    rq_activate_all_grippers(True)
    # end: URCap Program Node
  end
  $ 64 "zero_ftsensor()"
  zero_ftsensor()
  $ 65 "EXTT"
  $ 66 "Set GRP_3F_Enable=Off"
  set_standard_digital_out(4, False)
  $ 67 "Set BarcodeTrigger=Off"
  set_standard_digital_out(6, False)
  $ 68 "Set GRP_3F_Decap=Off"
  set_standard_digital_out(3, False)
  $ 69 "Set GRP_3F_Cap=Off"
  set_standard_digital_out(2, False)
  $ 70 "Set GRP_3F_Open=Off"
  set_standard_digital_out(5, False)
  $ 71 "PSE_T≔get_tool_free_pose(dir=[0,0,0.150], move_in_base_frame=True)"
  global PSE_T=get_tool_free_pose(dir=[0,0,0.150], move_in_base_frame=True)
  $ 72 "If is_reachable(Base_const, [PSE_T])"
  if (is_reachable(p[0.0,0.0,0.0,0.0,0.0,0.0], [PSE_T])):
    $ 73 "MoveL"
    $ 74 "PSE_T" "breakAfter"
    movel(PSE_T, a=1.2, v=0.15)
  end
  $ 76 "powder dispensing variable init"
  $ 77 "Start_thread≔ False "
  global Start_thread=  False
  $ 78 "vib_thread≔ False "
  global vib_thread=  False
  $ 79 "QR assignment init"
  $ 80 "d_cc≔0.06"
  global d_cc=0.06
  $ 81 "W_EMPTY≔50.131"
  global W_EMPTY=50.131
  $ 82 "kp≔0.0015"
  global kp=0.0015
  $ 83 "ki≔0.0001"
  global ki=0.0001
  $ 84 "kd≔0.01"
  global kd=0.01
  $ 85 "dt≔0.03"
  global dt=0.03
  $ 86 "Integral_error≔0"
  global Integral_error=0
  $ 87 "current_error≔0"
  global current_error=0
  $ 88 "previous_error≔0"
  global previous_error=0
  $ 89 "tilt_increment≔0"
  global tilt_increment=0
  $ 90 "tilt_angle≔0"
  global tilt_angle=0
  $ 91 "diff≔0"
  global diff=0
  $ 92 "current_pose≔get_actual_tcp_pose()"
  global current_pose= get_actual_tcp_pose ()
  $ 93 "Relative_trans≔p[0, 0, -0.035, 0, 0, 0]"
  global Relative_trans=p[0, 0, -0.035, 0, 0, 0]
  $ 97 "tilt_init_reference()"
  tilt_init_reference()
  $ 98 "switch_spat_M≔ True "
  global switch_spat_M=  True
  $ 99 "switch_spat_S≔ True "
  global switch_spat_S=  True
  $ 100 "switch_spat_F_M≔ True "
  global switch_spat_F_M=  True
  $ 101 "switch_spat_F_S≔ True "
  global switch_spat_F_S=  True
  $ 102 "last_scale≔0"
  global last_scale=0
  $ 775 "Thread_1"
  thread Thread_1():
    while (True):
      $ 776 "If Start_thread≟ True "
      if (Start_thread ==   True  ):
        $ 777 "weight_value≔get_weight()"
        global weight_value=get_weight()
        $ 778 "Wait: 0.1"
        sleep(0.1)
        $ 779 "sync()"
        sync()
      end
      $ 780 "sync()"
      sync()
    end
  end
  threadId_Thread_1 = run Thread_1()
  $ 781 "Thread_2"
  thread Thread_2():
    while (True):
      $ 782 "Loop vib_thread≟ True "
      thread Thread_while_782():
        while (True):
          $ 783 "diff≔target_weight-weight_value"
          global diff=target_weight-weight_value
          $ 784 "If diff>0.02 and spatula≠'spatula_flat_S'"
          global thread_flag_784=0
          thread Thread_if_784():
            $ 786 "Set AO[0]=4.0"
            set_standard_analog_out(0, 0.4)
            thread_flag_784 = 1
          end
          if (diff>0.02  and  spatula != "spatula_flat_S"):
            global thread_handler_784=run Thread_if_784()
            while (thread_flag_784 == 0):
              if not(diff>0.02  and  spatula != "spatula_flat_S"):
                kill thread_handler_784
                thread_flag_784 = 2
              else:
                sync()
              end
            end
          else:
            thread_flag_784 = 2
          end
          if (thread_flag_784 == 2):
            $ 787 "ElseIf diff>0.02 and spatula≟'spatula_flat_S'"
            if (diff>0.02 and spatula == "spatula_flat_S"):
              $ 788 "vibration_3()"
              vibration_3()
            else:
              $ 789 "ElseIf diff≤0.03"
              global thread_flag_789=0
              thread Thread_if_789():
                $ 790 "vibration_2()"
                vibration_2()
                thread_flag_789 = 1
              end
              if (diff <= 0.03):
                global thread_handler_789=run Thread_if_789()
                while (thread_flag_789 == 0):
                  if not(diff <= 0.03):
                    kill thread_handler_789
                    thread_flag_789 = 2
                  else:
                    sync()
                  end
                end
              else:
                thread_flag_789 = 2
              end
              if (thread_flag_789 == 2):
                $ 795 "Else" "noBreak"
                $ 796 "Set AO[0]=0.0"
                set_standard_analog_out(0, 0.0)
              end
            end
          end
        end
      end
      if (vib_thread ==   True  ):
        global thread_handler_782=run Thread_while_782()
        while (vib_thread ==   True  ):
          sync()
        end
        kill thread_handler_782
      end
      $ 797 "sync()"
      sync()
    end
  end
  threadId_Thread_2 = run Thread_2()
  while (True):
    $ 103 "Robot Program"
    $ 104 "MAIN"
    $ 105 "command_manager(external_control='uGO', cond_suspend=(ITM_Manipulated and AMR_AtTarget and AMR_Charging and AMR_Battery<40), cond_unsuspend=(AMR_Battery≟60))"
    command_manager(external_control="uGO", cond_suspend=(ITM_Manipulated  and  AMR_AtTarget  and  AMR_Charging  and  AMR_Battery<40), cond_unsuspend=(AMR_Battery == 60))
    $ 106 "log_state(STATE_Info)"
    log_state(STATE_Info)
    $ 107 "Switch STATE"
    switch_1 = STATE
    $ 108 "Case 1"
    if (1 == switch_1):
      $ 109 "Stopping"
      $ 110 "STATE_Info≔'Stopping'"
      global STATE_Info="Stopping"
      $ 111 "end_freedrive_mode()"
      end_freedrive_mode()
      $ 112 "Set"
      set_tcp(p[0.0,0.0,0.161,3.1415,0.0,0.0])
      $ 113 "PSE_T≔get_tool_free_pose(dir=[0,0,0.150], move_in_base_frame=True)"
      global PSE_T=get_tool_free_pose(dir=[0,0,0.150], move_in_base_frame=True)
      $ 114 "If is_reachable(Base_const, [PSE_T])"
      if (is_reachable(p[0.0,0.0,0.0,0.0,0.0,0.0], [PSE_T])):
        $ 115 "MoveL"
        $ 116 "PSE_T" "breakAfter"
        movel(PSE_T, a=1.2, v=0.15)
      end
      $ 117 "do_transition(keep_rxry=OBJ_Picked, r=0)"
      do_transition(keep_rxry=OBJ_Picked, r=0)
      $ 126 "Call Sub_AMR_MiR_V3"
      Sub_AMR_MiR_V3()
      $ 127 "If stopping() and AMR_Done"
      if (stopping()  and  AMR_Done):
        $ 128 "STATE≔2"
        global STATE=2
        $ 129 "ugo_update_outputs()"
        ugo_update_outputs()
      end
    elif (2 == switch_1):
      $ 130 "Case 2"
      $ 131 "Stopped"
      $ 132 "STATE_Info≔'Stopped'"
      global STATE_Info="Stopped"
      $ 133 "Call Sub_AMR_MiR_V3"
      Sub_AMR_MiR_V3()
      $ 134 "If CMD_Reset  or PB_Start"
      if (CMD_Reset   or  get_standard_digital_in(0)):
        $ 135 "STATE≔3"
        global STATE=3
        $ 136 "ugo_update_outputs()"
        ugo_update_outputs()
      end
    elif (3 == switch_1):
      $ 137 "Case 3"
      $ 138 " Resetting"
      $ 139 "STATE_Info≔'Resetting'"
      global STATE_Info="Resetting"
      $ 140 "uML"
      $ 141 "reset_error()"
      reset_error()
      $ 142 "reset_warning()"
      reset_warning()
      $ 143 "PROCESS_Step≔0"
      global PROCESS_Step=0
      $ 144 "PROCESS_Info≔''"
      global PROCESS_Info=""
      $ 145 "ARM_Referenced≔ False "
      global ARM_Referenced=  False
      $ 146 "WRK_Done≔ False "
      global WRK_Done=  False
      $ 147 "ITM_Prepared≔ False "
      global ITM_Prepared=  False
      $ 148 "ITM_Manipulated≔ False "
      global ITM_Manipulated=  False
      $ 149 "STP≔0"
      global STP=0
      $ 150 "Action≔0"
      global Action=0
      $ 151 "Action_Info≔''"
      global Action_Info=""
      $ 152 "ITM_ID≔0"
      global ITM_ID=0
      $ 153 "JIG≔0"
      global JIG=0
      $ 154 "JIG_Slot≔0"
      global JIG_Slot=0
      $ 155 "Task_info≔''"
      global Task_info=""
      $ 156 "Set"
      set_tcp(p[0.0,0.0,0.161,3.1415,0.0,0.0])
      $ 157 "App"
      $ 158 "'ADD APPLICATION SPECIFIC COMMANDS'"
      # 'ADD APPLICATION SPECIFIC COMMANDS'
      $ 159 "OBJ_Type≔0"
      global OBJ_Type=0
      $ 160 "OBJ_Nbr≔0"
      global OBJ_Nbr=0
      $ 161 "If CNT_Rack_Output≥50"
      if (CNT_Rack_Output >= 50):
        $ 162 "CNT_Rack_Output≔0"
        global CNT_Rack_Output=0
      end
      $ 163 "TASK≔struct(ID=0, NAVI=struct(target=0, footprint=0, protectiveOff=0, dock=0), WORK=struct(ITM_ID_Src=0, JIG_ID_Src=0, OBJ_Nbr_Src=0, ACT_Src=0, ITM_ID_Tgt=0, JIG_ID_Tgt=0, OBJ_Nbr_Tgt=0, ACT_Tgt=0, OBJ_Type=0))"
      global TASK=struct(ID=0, NAVI=struct(target=0, footprint=0, protectiveOff=0, dock=0), WORK=struct(ITM_ID_Src=0, JIG_ID_Src=0, OBJ_Nbr_Src=0, ACT_Src=0, ITM_ID_Tgt=0, JIG_ID_Tgt=0, OBJ_Nbr_Tgt=0, ACT_Tgt=0, OBJ_Type=0))
      $ 164 "Call Sub_AMR_MiR_V3"
      Sub_AMR_MiR_V3()
      $ 165 "If resetting() and AMR_Done"
      if (resetting()  and  AMR_Done):
        $ 166 "STATE≔4"
        global STATE=4
        $ 167 "ugo_update_outputs()"
        ugo_update_outputs()
      end
    elif (4 == switch_1):
      $ 168 "Case 4"
      $ 169 "Idle"
      $ 170 "STATE_Info≔'Idle'"
      global STATE_Info="Idle"
      $ 171 "If CMD_Start"
      if (CMD_Start):
        $ 172 "STATE≔5"
        global STATE=5
        $ 173 "ugo_update_outputs()"
        ugo_update_outputs()
      end
    elif (5 == switch_1):
      $ 174 "Case 5"
      $ 175 "Starting"
      $ 176 "STATE_Info≔'Starting'"
      global STATE_Info="Starting"
      $ 177 "'ADD COMMANDS WHAT TO START WITH'"
      # 'ADD COMMANDS WHAT TO START WITH'
      $ 178 "Call Sub_AMR_MiR_V3"
      Sub_AMR_MiR_V3()
      $ 179 "get ugo data"
      $ 180 "Assign Tasks"
      $ 181 "TASK.ID = ugo_get_task()"
      TASK.ID = ugo_get_task()
      $ 182 "If TASK.ID≟1"
      if (TASK.ID == 1):
        $ 183 "Task_info≔'Charge'"
        global Task_info="Charge"
        $ 184 "Parameters"
        $ 185 "AMR_PosTarget≔1"
        global AMR_PosTarget=1
      else:
        $ 186 "ElseIf TASK.ID≟9"
        if (TASK.ID == 9):
          $ 187 "'Pick Sarstedt Rack from Variable source'"
          # 'Pick Sarstedt Rack from Variable source'
          $ 188 "Task_info≔'Navigate to Target'"
          global Task_info="Navigate to Target"
          $ 189 "Parameters"
          $ 190 "AMR_PosTarget≔UGO.read_input('00','ITM_ID')"
          global AMR_PosTarget=UGO.read_input("00","ITM_ID")
        else:
          $ 191 "ElseIf TASK.ID≟49"
          if (TASK.ID == 49):
            $ 192 "Task_info≔'Pick Containers'"
            global Task_info="Pick Containers"
            $ 193 "Parameters"
            $ 194 "ITM_ID≔1"
            global ITM_ID=1
            $ 195 "OBJ_Type≔6"
            global OBJ_Type=6
            $ 196 "JIG≔15"
            global JIG=15
            $ 197 "AMR_PosTarget≔3"
            global AMR_PosTarget=3
          else:
            $ 198 "ElseIf TASK.ID≟50"
            if (TASK.ID == 50):
              $ 199 "Task_info≔'Decap Containers'"
              global Task_info="Decap Containers"
              $ 200 "Parameters"
              $ 201 "ITM_ID≔1"
              global ITM_ID=1
              $ 202 "OBJ_Type≔6"
              global OBJ_Type=6
              $ 203 "JIG≔16"
              global JIG=16
              $ 204 "AMR_PosTarget≔5"
              global AMR_PosTarget=5
            else:
              $ 205 "ElseIf TASK.ID≟51"
              if (TASK.ID == 51):
                $ 206 "Task_info≔'Detect Spatula and transfer powder'"
                global Task_info="Detect Spatula and transfer powder"
                $ 207 "Parameters"
                $ 208 "ITM_ID≔1"
                global ITM_ID=1
                $ 209 "target_weight≔(UGO.read_input('00','Target_weight'))/1000"
                global target_weight=(UGO.read_input("00","Target_weight"))/1000
                $ 210 "OBJ_Type≔8"
                global OBJ_Type=8
                $ 211 "JIG≔16"
                global JIG=16
                $ 212 "AMR_PosTarget≔5"
                global AMR_PosTarget=5
              else:
                $ 213 "ElseIf TASK.ID≟52"
                if (TASK.ID == 52):
                  $ 214 "Task_info≔'Pick Powder'"
                  global Task_info="Pick Powder"
                  $ 215 "Parameters"
                  $ 216 "ITM_ID≔1"
                  global ITM_ID=1
                  $ 217 "OBJ_Type≔6"
                  global OBJ_Type=6
                  $ 218 "JIG≔15"
                  global JIG=15
                  $ 219 "AMR_PosTarget≔3"
                  global AMR_PosTarget=3
                else:
                  $ 220 "ElseIf TASK.ID≟53"
                  if (TASK.ID == 53):
                    $ 221 "Task_info≔'Decap Powder'"
                    global Task_info="Decap Powder"
                    $ 222 "Parameters"
                    $ 223 "ITM_ID≔1"
                    global ITM_ID=1
                    $ 224 "OBJ_Type≔6"
                    global OBJ_Type=6
                    $ 225 "JIG≔1"
                    global JIG=1
                    $ 226 "AMR_PosTarget≔5"
                    global AMR_PosTarget=5
                  else:
                    $ 227 "ElseIf TASK.ID≟54"
                    if (TASK.ID == 54):
                      $ 228 "Task_info≔'Empty and swap Powder container'"
                      global Task_info="Empty and swap Powder container"
                      $ 237 "Parameters"
                      $ 238 "ITM_ID≔1"
                      global ITM_ID=1
                      $ 240 "W_now≔(UGO.read_input('00','Container_weight'))/1000"
                      global W_now=(UGO.read_input("00","Container_weight"))/1000
                      $ 241 "Pow_name≔(UGO.read_input('00','Powder_name'))"
                      global Pow_name=(UGO.read_input("00","Powder_name"))
                      $ 242 "scooping_init()"
                      scooping_init()
                      $ 243 "target_weight≔W_now-W_EMPTY-(0.002*W_FULL)"
                      global target_weight=W_now-W_EMPTY-(0.002*W_FULL)
                      $ 244 "OBJ_Type≔6"
                      global OBJ_Type=6
                      $ 245 "JIG≔17"
                      global JIG=17
                      $ 246 "AMR_PosTarget≔5"
                      global AMR_PosTarget=5
                    else:
                      $ 247 "ElseIf TASK.ID≟55"
                      if (TASK.ID == 55):
                        $ 248 "Task_info≔'Place Powder'"
                        global Task_info="Place Powder"
                        $ 249 "Parameters"
                        $ 250 "ITM_ID≔1"
                        global ITM_ID=1
                        $ 251 "OBJ_Type≔6"
                        global OBJ_Type=6
                        $ 252 "JIG≔21"
                        global JIG=21
                        $ 253 "AMR_PosTarget≔5"
                        global AMR_PosTarget=5
                      else:
                        $ 254 "ElseIf TASK.ID≟56"
                        if (TASK.ID == 56):
                          $ 255 "Task_info≔'Dose Powder'"
                          global Task_info="Dose Powder"
                          $ 256 "Parameters"
                          $ 257 "ITM_ID≔1"
                          global ITM_ID=1
                          $ 258 "target_weight≔(UGO.read_input('00','Target_weight'))/1000"
                          global target_weight=(UGO.read_input("00","Target_weight"))/1000
                          $ 259 "W_now≔(UGO.read_input('00','Container_weight'))/1000"
                          global W_now=(UGO.read_input("00","Container_weight"))/1000
                          $ 261 "Pow_name≔(UGO.read_input('00','Powder_name'))"
                          global Pow_name=(UGO.read_input("00","Powder_name"))
                          $ 262 "OBJ_Type≔6"
                          global OBJ_Type=6
                          $ 263 "JIG≔17"
                          global JIG=17
                          $ 264 "AMR_PosTarget≔5"
                          global AMR_PosTarget=5
                        else:
                          $ 265 "ElseIf TASK.ID≟57"
                          if (TASK.ID == 57):
                            $ 266 "Task_info≔'Recipe Powder dosing'"
                            global Task_info="Recipe Powder dosing"
                            $ 267 "Parameters"
                            $ 268 "ITM_ID≔1"
                            global ITM_ID=1
                            $ 269 "Pow_A≔(UGO.read_input('00','PowderA'))"
                            global Pow_A=(UGO.read_input("00","PowderA"))
                            $ 270 "Pow_B≔(UGO.read_input('00','PowderB'))"
                            global Pow_B=(UGO.read_input("00","PowderB"))
                            $ 271 "Pow_C≔(UGO.read_input('00','PowderC'))"
                            global Pow_C=(UGO.read_input("00","PowderC"))
                            $ 272 "Total_weight≔(UGO.read_input('00','Total_weight'))/1000"
                            global Total_weight=(UGO.read_input("00","Total_weight"))/1000
                            $ 273 "Pow_A_percent≔(UGO.read_input('00','PowderA_percentage'))/100"
                            global Pow_A_percent=(UGO.read_input("00","PowderA_percentage"))/100
                            $ 274 "Pow_B_percent≔(UGO.read_input('00','PowderB_percentage'))/100"
                            global Pow_B_percent=(UGO.read_input("00","PowderB_percentage"))/100
                            $ 275 "Pow_C_percent≔(UGO.read_input('00','PowderC_percentage'))/100"
                            global Pow_C_percent=(UGO.read_input("00","PowderC_percentage"))/100
                            $ 276 "OBJ_Type≔6"
                            global OBJ_Type=6
                            $ 277 "JIG≔17"
                            global JIG=17
                            $ 278 "AMR_PosTarget≔5"
                            global AMR_PosTarget=5
                          else:
                            $ 279 "ElseIf TASK.ID≟58"
                            if (TASK.ID == 58):
                              $ 280 "Task_info≔'Pick Powder containers'"
                              global Task_info="Pick Powder containers"
                              $ 281 "Parameters"
                              $ 282 "ITM_ID≔1"
                              global ITM_ID=1
                              $ 283 "OBJ_Type≔6"
                              global OBJ_Type=6
                              $ 284 "JIG≔15"
                              global JIG=15
                              $ 285 "AMR_PosTarget≔3"
                              global AMR_PosTarget=3
                            else:
                              $ 286 "Else" "noBreak"
                              $ 287 "set_error(ERROR_WRONG_ORDER)"
                              set_error(ERROR_WRONG_ORDER)
                            end
                          end
                        end
                      end
                    end
                  end
                end
              end
            end
          end
        end
      end
      $ 288 "test ugo"
      $ 289 "Wait: 0.2"
      sleep(0.2)
      $ 290 "ugo_update_outputs()"
      ugo_update_outputs()
      $ 291 "If starting() and AMR_Done"
      if (starting()  and  AMR_Done):
        $ 292 "log_message(Task_info, 'New Task: ')"
        log_message(Task_info, "New Task: ")
        $ 293 "log_message(to_str(TASK.ID), 'Task_ID: ')"
        log_message(to_str(TASK.ID), "Task_ID: ")
        $ 294 "do_transition(keep_rxry=OBJ_Picked)"
        do_transition(keep_rxry=OBJ_Picked)
        $ 295 "STATE≔6"
        global STATE=6
        $ 296 "ugo_update_outputs()"
        ugo_update_outputs()
      end
    elif (6 == switch_1):
      $ 297 "Case 6"
      $ 298 "Execute"
      $ 299 "STATE_Info≔'Execute'"
      global STATE_Info="Execute"
      $ 300 "If  not CMD_Hold and not CMD_Suspend"
      global thread_flag_300=0
      thread Thread_if_300():
        $ 301 "Switch PROCESS_Step"
        switch_2 = PROCESS_Step
        $ 302 "Case 0"
        if (0 == switch_2):
          $ 303 "PROCESS_Info≔'process control'"
          global PROCESS_Info="process control"
          $ 304 "log_process(PROCESS_Info)"
          log_process(PROCESS_Info)
          $ 305 "process control"
          $ 306 "If  not AMR_AtTarget"
          if (  not  AMR_AtTarget):
            $ 307 "PROCESS_Step≔1"
            global PROCESS_Step=1
          else:
            $ 308 "ElseIf (( not ITM_Prepared and  not WRK_Done) or (ITM_Prepared and WRK_Done))"
            if (((  not  ITM_Prepared  and    not  WRK_Done)  or  (ITM_Prepared  and  WRK_Done))):
              $ 309 "PROCESS_Step≔2"
              global PROCESS_Step=2
            else:
              $ 310 "ElseIf  not WRK_Done"
              if (  not  WRK_Done):
                $ 311 "PROCESS_Step≔3"
                global PROCESS_Step=3
              else:
                $ 312 "Else" "noBreak"
                $ 313 "task finished"
                $ 314 "PROCESS_Info≔''"
                global PROCESS_Info=""
                $ 315 "STATE≔7"
                global STATE=7
                $ 316 "ugo_update_outputs()"
                ugo_update_outputs()
              end
            end
          end
        elif (1 == switch_2):
          $ 317 "Case 1"
          $ 318 "navigate"
          $ 319 "'MOVING THE uML'"
          # 'MOVING THE uML'
          $ 320 "PROCESS_Info≔'move to target'"
          global PROCESS_Info="move to target"
          $ 321 "log_process(PROCESS_Info)"
          log_process(PROCESS_Info)
          $ 322 "If TASK.ID≟1"
          if (TASK.ID == 1):
            $ 323 "Action≔51"
            global Action=51
          else:
            $ 324 "Else" "noBreak"
            $ 325 "Action≔52"
            global Action=52
          end
          $ 326 "Call Sub_AMR_MiR_V3"
          Sub_AMR_MiR_V3()
          $ 327 "If AMR_Done"
          if (AMR_Done):
            $ 328 "PROCESS_Step≔0"
            global PROCESS_Step=0
          end
        elif (2 == switch_2):
          $ 329 "Case 2"
          $ 330 "prepare"
          $ 331 "'THINGS THAT HAVE TO BE DONE ONCE IN A SEQUENCE,WORKFLOW'"
          # 'THINGS THAT HAVE TO BE DONE ONCE IN A SEQUENCE,WORKFLOW'
          $ 332 "PROCESS_Info≔'prepare for work'"
          global PROCESS_Info="prepare for work"
          $ 333 "log_process(PROCESS_Info)"
          log_process(PROCESS_Info)
          $ 334 "If TASK.WORK.ITM_ID_Src>1"
          if (TASK.WORK.ITM_ID_Src>1):
            $ 335 "ITM_ID≔TASK.WORK.ITM_ID_Src"
            global ITM_ID=TASK.WORK.ITM_ID_Src
          else:
            $ 336 "ElseIf TASK.WORK.ITM_ID_Tgt>1"
            if (TASK.WORK.ITM_ID_Tgt>1):
              $ 337 "ITM_ID≔TASK.WORK.ITM_ID_Tgt"
              global ITM_ID=TASK.WORK.ITM_ID_Tgt
            end
          end
          $ 338 "If  not ARM_Referenced and (ITM_ID≠0)"
          if (  not  ARM_Referenced  and  (ITM_ID != 0)):
            $ 339 "STP≔1"
            global STP=1
          else:
            $ 340 "ElseIf ARM_Referenced or (ITM_ID≟0)"
            if (ARM_Referenced  or  (ITM_ID == 0)):
              $ 341 "STP≔2"
              global STP=2
            end
          end
          $ 342 "Switch STP"
          switch_3 = STP
          $ 343 "Case 1"
          if (1 == switch_3):
            $ 344 "reference"
            $ 345 "STP_Info≔'reference at target position'"
            global STP_Info="reference at target position"
            $ 346 "log_step(STP_Info)"
            log_step(STP_Info)
            $ 347 "If ITM_ID≟1"
            if (ITM_ID == 1):
              $ 348 "CAM_Done≔ True "
              global CAM_Done=  True
            else:
              $ 349 "Else" "noBreak"
              $ 350 "Action≔131"
              global Action=131
              $ 351 "Call Sub_Vision_V18"
              Sub_Vision_V18()
            end
            $ 353 "If CAM_Done and  not ERROR.FLAG"
            if (CAM_Done  and    not  ERROR.FLAG):
              $ 354 "log_step('ARM referenced')"
              log_step("ARM referenced")
              $ 355 "ARM_Referenced≔ True "
              global ARM_Referenced=  True
            end
          elif (2 == switch_3):
            $ 356 "Case 2"
            $ 357 "manipulate"
            $ 358 "STP_Info≔'manipulate item'"
            global STP_Info="manipulate item"
            $ 359 "log_step(STP_Info)"
            log_step(STP_Info)
            $ 360 "'In case pressing button is needed'"
            # 'In case pressing button is needed'
            $ 361 "If found_in_list(ITM_ID, ITM_ID_List)"
            if (found_in_list(ITM_ID, ITM_ID_List)):
              $ 362 "Switch ITM_ID"
              switch_4 = ITM_ID
              $ 363 "Case 0"
              if (0 == switch_4):
                $ 364 "ITM_Manipulated≔ not ITM_Manipulated"
                global ITM_Manipulated=  not  ITM_Manipulated
              elif (1 == switch_4):
                $ 365 "Case 1"
                $ 366 "ITM_Manipulated≔ not ITM_Manipulated"
                global ITM_Manipulated=  not  ITM_Manipulated
              elif (2 == switch_4):
                $ 367 "Case 2"
              else:
                $ 377 "Default Case"
                $ 378 "ITM_Manipulated≔ not ITM_Manipulated"
                global ITM_Manipulated=  not  ITM_Manipulated
              end
            end
          end
          $ 379 "ITM_Prepared≔(ITM_Manipulated or  not found_in_list(ITM_ID, ITM_ID_List)) and (ARM_Referenced or ITM_ID≟0) and  not WRK_Done"
          global ITM_Prepared=(ITM_Manipulated  or    not  found_in_list(ITM_ID, ITM_ID_List))  and  (ARM_Referenced  or  ITM_ID == 0)  and    not  WRK_Done
          $ 380 "STP≔0"
          global STP=0
          $ 381 "STP_Info≔''"
          global STP_Info=""
          $ 382 "PROCESS_Step≔0"
          global PROCESS_Step=0
        elif (3 == switch_2):
          $ 383 "Case 3"
          $ 384 "work"
          $ 385 "'ADD EVERY MACHINE, OBJECT, STATION TO WORK ON'"
          # 'ADD EVERY MACHINE, OBJECT, STATION TO WORK ON'
          $ 386 "Switch ITM_ID"
          switch_3 = ITM_ID
          $ 387 "Case 1"
          if (1 == switch_3):
            $ 388 "uLM"
            $ 389 "If TASK.ID≟12"
            if (TASK.ID == 12):
              $ 390 "fill racks"
              $ 391 "Action≔151"
              global Action=151
              $ 392 "Call Sub_Vision_V18"
              Sub_Vision_V18()
              $ 393 "If  not ERROR.FLAG"
              if (  not  ERROR.FLAG):
                $ 394 "Actions for the task"
                $ 395 "Action≔1"
                global Action=1
                $ 396 "JIG≔2"
                global JIG=2
                $ 397 "JIG_Slot≔CAM_Result[0]"
                global JIG_Slot=CAM_Result[0]
                $ 398 "OBJ_Nbr≔CAM_Result[0]"
                global OBJ_Nbr=CAM_Result[0]
                $ 399 "OBJ_Type≔2"
                global OBJ_Type=2
                $ 400 "Call Sub_Action_V4"
                Sub_Action_V4()
                $ 401 "If OBJ_Picked"
                if (OBJ_Picked):
                  $ 402 "CAM_Result.remove(0)"
                  CAM_Result.remove(0)
                  $ 403 "PRC_TubCounter≔PRC_TubCounter+1"
                  global PRC_TubCounter=PRC_TubCounter+1
                  $ 404 "If PRC_TubCounter%4≟0"
                  if (PRC_TubCounter%4 == 0):
                    $ 405 "JIG_Slot≔4"
                    global JIG_Slot=4
                  else:
                    $ 406 "Else" "noBreak"
                    $ 407 "JIG_Slot≔PRC_TubCounter%4"
                    global JIG_Slot=PRC_TubCounter%4
                  end
                  $ 408 "OBJ_Nbr≔ceil(PRC_TubCounter/4)"
                  global OBJ_Nbr=ceil(PRC_TubCounter/4)
                  $ 409 "Action≔2"
                  global Action=2
                  $ 410 "JIG≔4"
                  global JIG=4
                  $ 411 "Call Sub_Action_V4"
                  Sub_Action_V4()
                  $ 412 "Action≔151"
                  global Action=151
                  $ 413 "Call Sub_Vision_V18"
                  Sub_Vision_V18()
                end
              end
              $ 414 "If (CAM_Captures≥CAM_PRM_Retries) or (PRC_TubCounter≥32)"
              if ((CAM_Captures >= CAM_PRM_Retries)  or  (PRC_TubCounter >= 32)):
                $ 415 "PROCESS_Step≔0"
                global PROCESS_Step=0
                $ 416 "WRK_Done≔ True "
                global WRK_Done=  True
              end
            else:
              $ 417 "ElseIf TASK.ID≟49"
              if (TASK.ID == 49):
                $ 418 "Pick Powder container"
                $ 419 "Action≔131"
                global Action=131
                $ 420 "Call Sub_Vision_V18"
                Sub_Vision_V18()
                $ 421 "Action≔35"
                global Action=35
                $ 422 "Call Sub_Action_V4"
                Sub_Action_V4()
                $ 423 "PROCESS_Step≔0"
                global PROCESS_Step=0
                $ 424 "WRK_Done≔ True "
                global WRK_Done=  True
              else:
                $ 425 "ElseIf TASK.ID≟50"
                if (TASK.ID == 50):
                  $ 426 "Decap containers"
                  $ 427 "Action≔36"
                  global Action=36
                  $ 428 "Call Sub_Action_V4"
                  Sub_Action_V4()
                  $ 429 "PROCESS_Step≔0"
                  global PROCESS_Step=0
                  $ 430 "WRK_Done≔ True "
                  global WRK_Done=  True
                else:
                  $ 431 "ElseIf TASK.ID≟51"
                  if (TASK.ID == 51):
                    $ 432 "Detect Spatula and transfer powder"
                    $ 433 "Action≔131"
                    global Action=131
                    $ 434 "Call Sub_Vision_V18"
                    Sub_Vision_V18()
                    $ 435 "Action≔37"
                    global Action=37
                    $ 436 "Call Sub_Action_V4"
                    Sub_Action_V4()
                    $ 437 "PROCESS_Step≔0"
                    global PROCESS_Step=0
                    $ 438 "WRK_Done≔ True "
                    global WRK_Done=  True
                  else:
                    $ 439 "ElseIf TASK.ID≟52"
                    if (TASK.ID == 52):
                      $ 440 "Pick Powder container"
                      $ 441 "Action≔131"
                      global Action=131
                      $ 442 "Call Sub_Vision_V18"
                      Sub_Vision_V18()
                      $ 443 "Action≔39"
                      global Action=39
                      $ 444 "Call Sub_Action_V4"
                      Sub_Action_V4()
                      $ 445 "PROCESS_Step≔0"
                      global PROCESS_Step=0
                      $ 446 "WRK_Done≔ True "
                      global WRK_Done=  True
                    else:
                      $ 447 "ElseIf TASK.ID≟53"
                      if (TASK.ID == 53):
                        $ 448 "Decap containerA"
                        $ 449 "Action≔40"
                        global Action=40
                        $ 450 "Call Sub_Action_V4"
                        Sub_Action_V4()
                        $ 451 "PROCESS_Step≔0"
                        global PROCESS_Step=0
                        $ 452 "WRK_Done≔ True "
                        global WRK_Done=  True
                      else:
                        $ 453 "ElseIf TASK.ID≟55"
                        if (TASK.ID == 55):
                          $ 454 "Place Powder"
                          $ 455 "Action≔131"
                          global Action=131
                          $ 456 "Call Sub_Vision_V18"
                          Sub_Vision_V18()
                          $ 457 "Action≔41"
                          global Action=41
                          $ 458 "Call Sub_Action_V4"
                          Sub_Action_V4()
                          $ 459 "PROCESS_Step≔0"
                          global PROCESS_Step=0
                          $ 460 "WRK_Done≔ True "
                          global WRK_Done=  True
                        else:
                          $ 461 "ElseIf TASK.ID≟54"
                          if (TASK.ID == 54):
                            $ 462 "Empty and swap container"
                            $ 463 "Action≔131"
                            global Action=131
                            $ 464 "Call Sub_Vision_V18"
                            Sub_Vision_V18()
                            $ 465 "Action≔42"
                            global Action=42
                            $ 466 "Call Sub_Action_V4"
                            Sub_Action_V4()
                            $ 467 "PROCESS_Step≔0"
                            global PROCESS_Step=0
                            $ 468 "WRK_Done≔ True "
                            global WRK_Done=  True
                          else:
                            $ 469 "ElseIf TASK.ID≟56"
                            if (TASK.ID == 56):
                              $ 470 "Dispense Powder"
                              $ 471 "Action≔131"
                              global Action=131
                              $ 472 "Call Sub_Vision_V18"
                              Sub_Vision_V18()
                              $ 473 "Action≔43"
                              global Action=43
                              $ 474 "Call Sub_Action_V4"
                              Sub_Action_V4()
                              $ 475 "PROCESS_Step≔0"
                              global PROCESS_Step=0
                              $ 476 "WRK_Done≔ True "
                              global WRK_Done=  True
                            else:
                              $ 477 "ElseIf TASK.ID≟57"
                              if (TASK.ID == 57):
                                $ 478 "Recipe Dosing"
                                $ 479 "Action≔48"
                                global Action=48
                                $ 480 "Call Sub_Action_V4"
                                Sub_Action_V4()
                                $ 481 "recipe_init(Pow_A, Pow_B, Pow_C, Total_weight, Pow_A_percent, Pow_B_percent, Pow_C_percent)"
                                recipe_init(Pow_A, Pow_B, Pow_C, Total_weight, Pow_A_percent, Pow_B_percent, Pow_C_percent)
                                $ 482 "Loop recipe_next()≟ True "
                                while (recipe_next() ==   True  ):
                                  $ 483 "Action≔44"
                                  global Action=44
                                  $ 484 "Call Sub_Action_V4"
                                  Sub_Action_V4()
                                  $ 485 "JIG≔21"
                                  global JIG=21
                                  $ 486 "Action≔131"
                                  global Action=131
                                  $ 487 "Call Sub_Vision_V18"
                                  Sub_Vision_V18()
                                  $ 488 "Action≔45"
                                  global Action=45
                                  $ 489 "Call Sub_Action_V4"
                                  Sub_Action_V4()
                                  $ 490 "dosing_start()"
                                  dosing_start()
                                  $ 491 "JIG≔17"
                                  global JIG=17
                                  $ 492 "Action≔131"
                                  global Action=131
                                  $ 493 "Call Sub_Vision_V18"
                                  Sub_Vision_V18()
                                  $ 494 "Action≔46"
                                  global Action=46
                                  $ 495 "Call Sub_Action_V4"
                                  Sub_Action_V4()
                                  $ 496 "dosing_end()"
                                  dosing_end()
                                end
                                $ 497 "PROCESS_Step≔0"
                                global PROCESS_Step=0
                                $ 498 "WRK_Done≔ True "
                                global WRK_Done=  True
                              else:
                                $ 499 "ElseIf TASK.ID≟58"
                                if (TASK.ID == 58):
                                  $ 500 "Pick Powder containers"
                                  $ 501 "Num_cont_picked≔0"
                                  global Num_cont_picked=0
                                  $ 502 "powder_position≔'Position1'"
                                  global powder_position="Position1"
                                  $ 503 "Loop Num_cont_picked<3"
                                  while (Num_cont_picked<3):
                                    $ 504 "Action≔131"
                                    global Action=131
                                    $ 505 "Call Sub_Vision_V18"
                                    Sub_Vision_V18()
                                    $ 506 "Action≔47"
                                    global Action=47
                                    $ 507 "Call Sub_Action_V4"
                                    Sub_Action_V4()
                                  end
                                  $ 508 "PROCESS_Step≔0"
                                  global PROCESS_Step=0
                                  $ 509 "WRK_Done≔ True "
                                  global WRK_Done=  True
                                end
                              end
                            end
                          end
                        end
                      end
                    end
                  end
                end
              end
            end
          elif (2 == switch_3):
            $ 510 "Case 2"
          elif (5 == switch_3):
            $ 552 "Case 5"
          elif (20 == switch_3):
            $ 560 "Case 20"
          elif (43 == switch_3):
            $ 622 "Case 43"
          else:
            $ 630 "Default Case"
            $ 631 "WRK_Done≔ True "
            global WRK_Done=  True
            $ 632 "PROCESS_Step≔0"
            global PROCESS_Step=0
          end
        end
        thread_flag_300 = 1
      end
      if (  not  CMD_Hold and not CMD_Suspend):
        global thread_handler_300=run Thread_if_300()
        while (thread_flag_300 == 0):
          if not(  not  CMD_Hold and not CMD_Suspend):
            kill thread_handler_300
            thread_flag_300 = 2
          else:
            sync()
          end
        end
      else:
        thread_flag_300 = 2
      end
      $ 633 "If CMD_Hold"
      if (CMD_Hold):
        $ 634 "STATE≔9"
        global STATE=9
        $ 635 "ugo_update_outputs()"
        ugo_update_outputs()
      else:
        $ 636 "ElseIf CMD_Suspend"
        if (CMD_Suspend):
          $ 637 "STATE≔12"
          global STATE=12
          $ 638 "ugo_update_outputs()"
          ugo_update_outputs()
        end
      end
    elif (7 == switch_1):
      $ 639 "Case 7"
      $ 640 "Completing"
      $ 641 "STATE_Info≔'Completing'"
      global STATE_Info="Completing"
      $ 642 "'ADD COMMANDS FOR COMPLETING THE PROCESS'"
      # 'ADD COMMANDS FOR COMPLETING THE PROCESS'
      $ 643 "do_transition(keep_rxry=OBJ_Picked)"
      do_transition(keep_rxry=OBJ_Picked)
      $ 644 "Call Sub_AMR_MiR_V3"
      Sub_AMR_MiR_V3()
      $ 645 "If completing() and AMR_Done"
      if (completing()  and  AMR_Done):
        $ 646 "STATE≔8"
        global STATE=8
        $ 647 "ugo_update_outputs()"
        ugo_update_outputs()
      end
    elif (8 == switch_1):
      $ 648 "Case 8"
      $ 649 "Complete"
      $ 650 "STATE_Info≔'Complete'"
      global STATE_Info="Complete"
      $ 651 "If CMD_Reset"
      if (CMD_Reset):
        $ 652 "STATE≔3"
        global STATE=3
        $ 653 "ugo_update_outputs()"
        ugo_update_outputs()
      end
    elif (9 == switch_1):
      $ 654 "Case 9"
      $ 655 "Holding"
      $ 656 "STATE_Info≔'Holding'"
      global STATE_Info="Holding"
      $ 657 "stopl(0.5)"
      stopl(0.5)
      $ 658 "Call Sub_AMR_MiR_V3"
      Sub_AMR_MiR_V3()
      $ 659 "If holding() and AMR_Done"
      if (holding()  and  AMR_Done):
        $ 660 "STATE≔10"
        global STATE=10
        $ 661 "ugo_update_outputs()"
        ugo_update_outputs()
      end
    elif (10 == switch_1):
      $ 662 "Case 10"
      $ 663 "Held"
      $ 664 "STATE_Info≔'Held'"
      global STATE_Info="Held"
      $ 665 "If CMD_Unhold"
      if (CMD_Unhold):
        $ 666 "end_freedrive_mode()"
        end_freedrive_mode()
        $ 667 "STATE≔11"
        global STATE=11
        $ 668 "ugo_update_outputs()"
        ugo_update_outputs()
      else:
        $ 669 "ElseIf FNC_Freedrive"
        if (FNC_Freedrive):
          $ 670 "freedrive_mode()"
          freedrive_mode()
        else:
          $ 671 "Else" "noBreak"
          $ 672 "end_freedrive_mode()"
          end_freedrive_mode()
        end
      end
    elif (11 == switch_1):
      $ 673 "Case 11"
      $ 674 "Unholding"
      $ 675 "STATE_Info≔'Unholding'"
      global STATE_Info="Unholding"
      $ 676 "Clearing"
      $ 677 "Switch ERROR.ID"
      switch_2 = ERROR.ID
      $ 678 "Case 1002"
      if (1002 == switch_2):
        $ 679 "AMR_AtTarget≔ False "
        global AMR_AtTarget=  False
        $ 680 "ARM_Referenced≔ False "
        global ARM_Referenced=  False
        $ 681 "ITM_Prepared≔ False "
        global ITM_Prepared=  False
        $ 682 "PROCESS_Step≔1"
        global PROCESS_Step=1
      elif (2007 == switch_2):
        $ 683 "Case 2007"
        $ 684 "PROCESS_Step≔1"
        global PROCESS_Step=1
      end
      $ 685 "reset_error()"
      reset_error()
      $ 686 "reset_warning()"
      reset_warning()
      $ 687 "OBJ_Picked≔gripper_has_object()"
      global OBJ_Picked=gripper_has_object()
      $ 688 "Call Sub_AMR_MiR_V3"
      Sub_AMR_MiR_V3()
      $ 689 "If unholding() and AMR_Done"
      if (unholding()  and  AMR_Done):
        $ 690 "STATE≔6"
        global STATE=6
        $ 691 "ugo_update_outputs()"
        ugo_update_outputs()
      end
    elif (12 == switch_1):
      $ 692 "Case 12"
      $ 693 "Suspending"
      $ 694 "STATE_Info≔'Suspending'"
      global STATE_Info="Suspending"
      $ 695 "PROCESS_Info≔str_cat(PROCESS_Info, ' suspended')"
      global PROCESS_Info=str_cat(PROCESS_Info, " suspended")
      $ 696 "If suspending()"
      if (suspending()):
        $ 697 "STATE≔13"
        global STATE=13
        $ 698 "ugo_update_outputs()"
        ugo_update_outputs()
      end
    elif (13 == switch_1):
      $ 699 "Case 13"
      $ 700 "Suspended"
      $ 701 "STATE_Info≔'Suspended'"
      global STATE_Info="Suspended"
      $ 702 "Call Sub_AMR_MiR_V3"
      Sub_AMR_MiR_V3()
      $ 703 "If CMD_Unsuspend"
      if (CMD_Unsuspend):
        $ 704 "STATE≔14"
        global STATE=14
        $ 705 "ugo_update_outputs()"
        ugo_update_outputs()
      end
    elif (14 == switch_1):
      $ 706 "Case 14"
      $ 707 "Unsuspending"
      $ 708 "STATE_Info≔'Unsuspending'"
      global STATE_Info="Unsuspending"
      $ 709 "PROCESS_Step≔0"
      global PROCESS_Step=0
      $ 710 "If unsuspending()"
      if (unsuspending()):
        $ 711 "STATE≔6"
        global STATE=6
        $ 712 "ugo_update_outputs()"
        ugo_update_outputs()
      end
    elif (15 == switch_1):
      $ 713 "Case 15"
      $ 714 "Aborting"
      $ 715 "STATE_Info≔'Aborting'"
      global STATE_Info="Aborting"
      $ 716 "If aborting()"
      if (aborting()):
        $ 717 "STATE≔16"
        global STATE=16
        $ 718 "ugo_update_outputs()"
        ugo_update_outputs()
      end
    elif (16 == switch_1):
      $ 719 "Case 16"
      $ 720 "Aborted"
      $ 721 "STATE_Info≔'Aborted'"
      global STATE_Info="Aborted"
      $ 722 "If CMD_Clear"
      if (CMD_Clear):
        $ 723 "STATE≔17"
        global STATE=17
        $ 724 "ugo_update_outputs()"
        ugo_update_outputs()
      end
    elif (17 == switch_1):
      $ 725 "Case 17"
      $ 726 "Clearing"
      $ 727 "STATE_Info≔'Clearing'"
      global STATE_Info="Clearing"
      $ 728 "Clearing"
      $ 729 "reset_warning()"
      reset_warning()
      $ 730 "reset_error()"
      reset_error()
      $ 731 "If clearing()"
      if (clearing()):
        $ 732 "STATE≔2"
        global STATE=2
        $ 733 "ugo_update_outputs()"
        ugo_update_outputs()
      end
    end
    $ 734 "log_state(STATE_Info)"
    log_state(STATE_Info)
    $ 735 "log_warning(WARNING.MSG)"
    log_warning(WARNING.MSG)
    $ 736 "log_error(ERROR.MSG)"
    log_error(ERROR.MSG)
    $ 737 "Times"
    $ 738 "Switch STATE"
    switch_1 = STATE
    $ 739 "Case 1"
    if (1 == switch_1):
      $ 740 "TM_St_Stopping≔get_time(STATE_Times[STATE-1])"
      global TM_St_Stopping=get_time(STATE_Times[STATE-1])
    elif (2 == switch_1):
      $ 741 "Case 2"
      $ 742 "TM_St_Stopped≔get_time(STATE_Times[STATE-1])"
      global TM_St_Stopped=get_time(STATE_Times[STATE-1])
    elif (3 == switch_1):
      $ 743 "Case 3"
      $ 744 "TM_St_Resetting≔get_time(STATE_Times[STATE-1])"
      global TM_St_Resetting=get_time(STATE_Times[STATE-1])
    elif (4 == switch_1):
      $ 745 "Case 4"
      $ 746 "TM_St_Idle≔get_time(STATE_Times[STATE-1])"
      global TM_St_Idle=get_time(STATE_Times[STATE-1])
    elif (5 == switch_1):
      $ 747 "Case 5"
      $ 748 "TM_St_Starting≔get_time(STATE_Times[STATE-1])"
      global TM_St_Starting=get_time(STATE_Times[STATE-1])
    elif (6 == switch_1):
      $ 749 "Case 6"
      $ 750 "TM_St_Execute≔get_time(STATE_Times[STATE-1])"
      global TM_St_Execute=get_time(STATE_Times[STATE-1])
    elif (7 == switch_1):
      $ 751 "Case 7"
      $ 752 "TM_St_Completin≔get_time(STATE_Times[STATE-1])"
      global TM_St_Completin=get_time(STATE_Times[STATE-1])
    elif (8 == switch_1):
      $ 753 "Case 8"
      $ 754 "TM_St_Complete≔get_time(STATE_Times[STATE-1])"
      global TM_St_Complete=get_time(STATE_Times[STATE-1])
    elif (9 == switch_1):
      $ 755 "Case 9"
      $ 756 "TM_St_Holding≔get_time(STATE_Times[STATE-1])"
      global TM_St_Holding=get_time(STATE_Times[STATE-1])
    elif (10 == switch_1):
      $ 757 "Case 10"
      $ 758 "TM_St_Held≔get_time(STATE_Times[STATE-1])"
      global TM_St_Held=get_time(STATE_Times[STATE-1])
    elif (11 == switch_1):
      $ 759 "Case 11"
      $ 760 "TM_St_Unholding≔get_time(STATE_Times[STATE-1])"
      global TM_St_Unholding=get_time(STATE_Times[STATE-1])
    elif (12 == switch_1):
      $ 761 "Case 12"
      $ 762 "TM_St_Suspendin≔get_time(STATE_Times[STATE-1])"
      global TM_St_Suspendin=get_time(STATE_Times[STATE-1])
    elif (13 == switch_1):
      $ 763 "Case 13"
      $ 764 "TM_St_Suspended≔get_time(STATE_Times[STATE-1])"
      global TM_St_Suspended=get_time(STATE_Times[STATE-1])
    elif (14 == switch_1):
      $ 765 "Case 14"
      $ 766 "TM_St_Unsuspend≔get_time(STATE_Times[STATE-1])"
      global TM_St_Unsuspend=get_time(STATE_Times[STATE-1])
    elif (15 == switch_1):
      $ 767 "Case 15"
      $ 768 "TM_St_Aborting≔get_time(STATE_Times[STATE-1])"
      global TM_St_Aborting=get_time(STATE_Times[STATE-1])
    elif (16 == switch_1):
      $ 769 "Case 16"
      $ 770 "TM_St_Aborted≔get_time(STATE_Times[STATE-1])"
      global TM_St_Aborted=get_time(STATE_Times[STATE-1])
    elif (17 == switch_1):
      $ 771 "Case 17"
      $ 772 "TM_St_Clearing≔get_time(STATE_Times[STATE-1])"
      global TM_St_Clearing=get_time(STATE_Times[STATE-1])
    end
    $ 774 "Wait: 0.1"
    sleep(0.1)
  end
end
